FUNCTION VERSION
  (* Standard: 61499-1 *)
  (* Version 1.0, 2024-03-05, franz *)
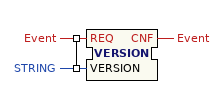
  EVENT_INPUT
    REQ WITH VERSION;
  END_EVENT
  EVENT_OUTPUT
    CNF;
  END_EVENT
  VAR_INPUT
    VERSION : STRING;
  END_VAR
  BODY IN ST:
FUNCTION VERSION
VAR_INPUT
	VERSION : STRING;
END_VAR
END_FUNCTION
  END_BODY
END_FUNCTION
